// SIMATIC S7-200 SMART project (STEP 7-Micro/WIN SMART), CPU SR30

SYMBOL_TABLE STATES
RUNNING_STATE    M4.0     // RUNNING STATE
ON_STATE         M0.0     // ON STATE
PROCESS          M0.1     // PROCESS START
X_AXIS_STATE     M0.2     // X_AXIS_STATE
Y_AXIS_STATE     M0.3     // Y_AXIS_STATE
GRIPPER_STATE    M0.4     // GRIPPER_STATE
PROGRAM_STARTED  M0.5     // PROGRAM STARTED
READY_STATE      M0.6     // READY_STATE
PAUSE_STATE      M0.7     // PAUSE_STATE
END_SYMBOL_TABLE

SYMBOL_TABLE STEPS
STEP_1_DONE      M1.0     // STEP_1_DONE
STEP_2_DONE      M1.1     // STEP_2_DONE
STEP_3_DONE      M1.2     // STEP_3_DONE
STEP_4_DONE      M1.3     // STEP_4_DONE
STEP_5_DONE      M1.4     // STEP_5_DONE
STEP_6_DONE      M1.5     // STEP_6_DONE
STEP_7_DONE      M1.6     // STEP_7_DONE
STEP_8_DONE      M1.7     // STEP_8_DONE
END_SYMBOL_TABLE

SYMBOL_TABLE HMI INPUTSS
HMI_START        M2.0     // HMI_START
HMI_PAUSE        M2.1     // HMI_PAUSE
HMI_STOP         M2.2     // HMI_STOP
HMI_E_STOP       M2.3     // HMI_E_STOP
END_SYMBOL_TABLE

SYMBOL_TABLE MASTER INPUTS
MASTER_STOP      V202.5   // MASTER_STOP
MASTER_START     V201.5   // MASTER_START
MASTER_RESET     V203.5   // MASTER_RESET
COMMUNCATION     M6.0     // COMMUNCATION
END_SYMBOL_TABLE

ORGANIZATION_BLOCK MAIN:OB1
TITLE=Program Comments
BEGIN
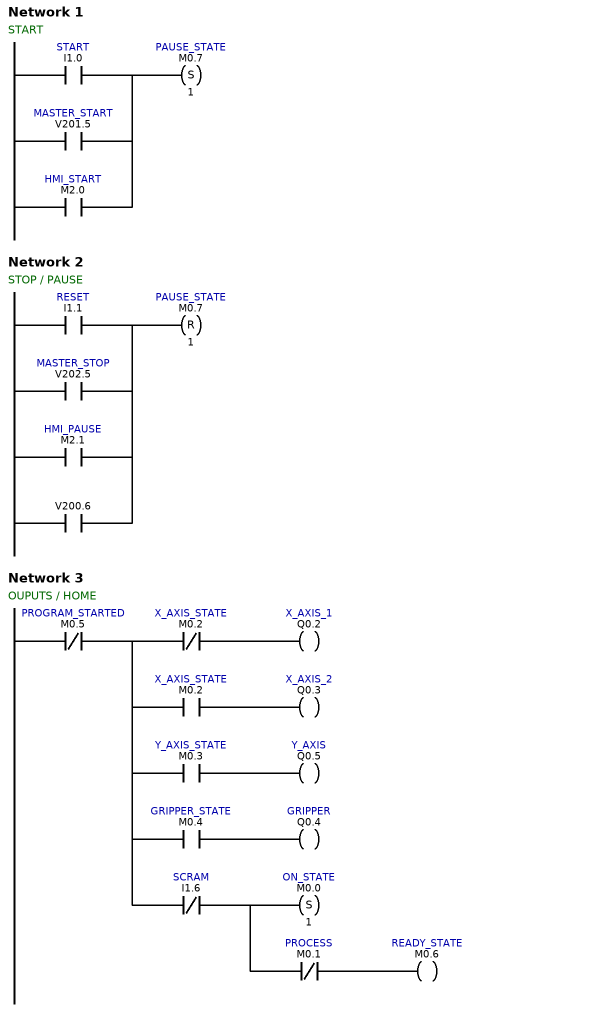
Network 1
// START
LD     START:I1.0
O      MASTER_START:V201.5
O      HMI_START:M2.0
S      PAUSE_STATE:M0.7, 1
Network 2
// STOP / PAUSE
LD     RESET:I1.1
O      MASTER_STOP:V202.5
O      HMI_PAUSE:M2.1
O      V200.6
R      PAUSE_STATE:M0.7, 1
Network 3
// OUPUTS / HOME
LDN    PROGRAM_STARTED:M0.5
LPS
AN     X_AXIS_STATE:M0.2
=      X_AXIS_1:Q0.2
LRD
A      X_AXIS_STATE:M0.2
=      X_AXIS_2:Q0.3
LRD
A      Y_AXIS_STATE:M0.3
=      Y_AXIS:Q0.5
LRD
A      GRIPPER_STATE:M0.4
=      GRIPPER:Q0.4
LPP
AN     SCRAM:I1.6
S      ON_STATE:M0.0, 1
AN     PROCESS:M0.1
=      READY_STATE:M0.6
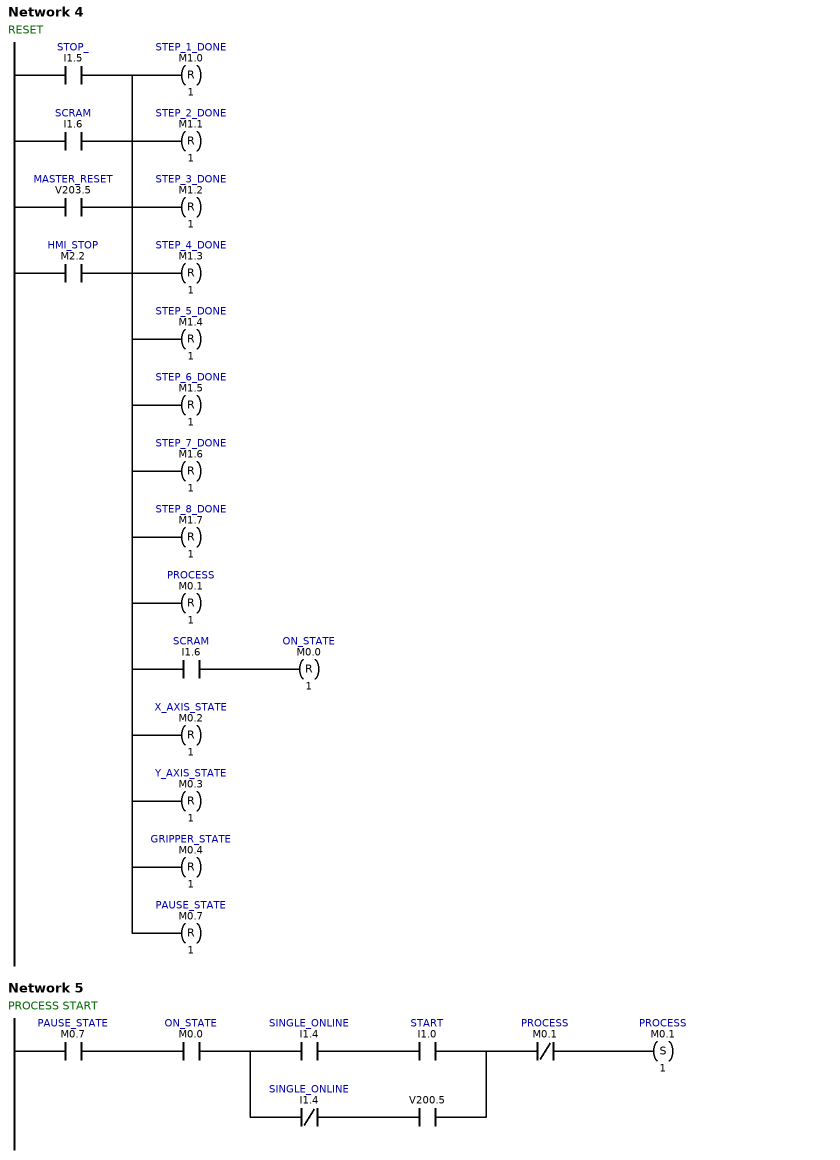
Network 4
// RESET 
LD     STOP_:I1.5
O      SCRAM:I1.6
O      MASTER_RESET:V203.5
O      HMI_STOP:M2.2
LPS
R      STEP_1_DONE:M1.0, 1
R      STEP_2_DONE:M1.1, 1
R      STEP_3_DONE:M1.2, 1
R      STEP_4_DONE:M1.3, 1
R      STEP_5_DONE:M1.4, 1
R      STEP_6_DONE:M1.5, 1
R      STEP_7_DONE:M1.6, 1
R      STEP_8_DONE:M1.7, 1
R      PROCESS:M0.1, 1
A      SCRAM:I1.6
R      ON_STATE:M0.0, 1
LRD
R      X_AXIS_STATE:M0.2, 1
LRD
R      Y_AXIS_STATE:M0.3, 1
LRD
R      GRIPPER_STATE:M0.4, 1
LPP
R      PAUSE_STATE:M0.7, 1
Network 5
// PROCESS START
LD     PAUSE_STATE:M0.7
A      ON_STATE:M0.0
LD     SINGLE_ONLINE:I1.4
A      START:I1.0
LDN    SINGLE_ONLINE:I1.4
A      V200.5
OLD
ALD
AN     PROCESS:M0.1
S      PROCESS:M0.1, 1
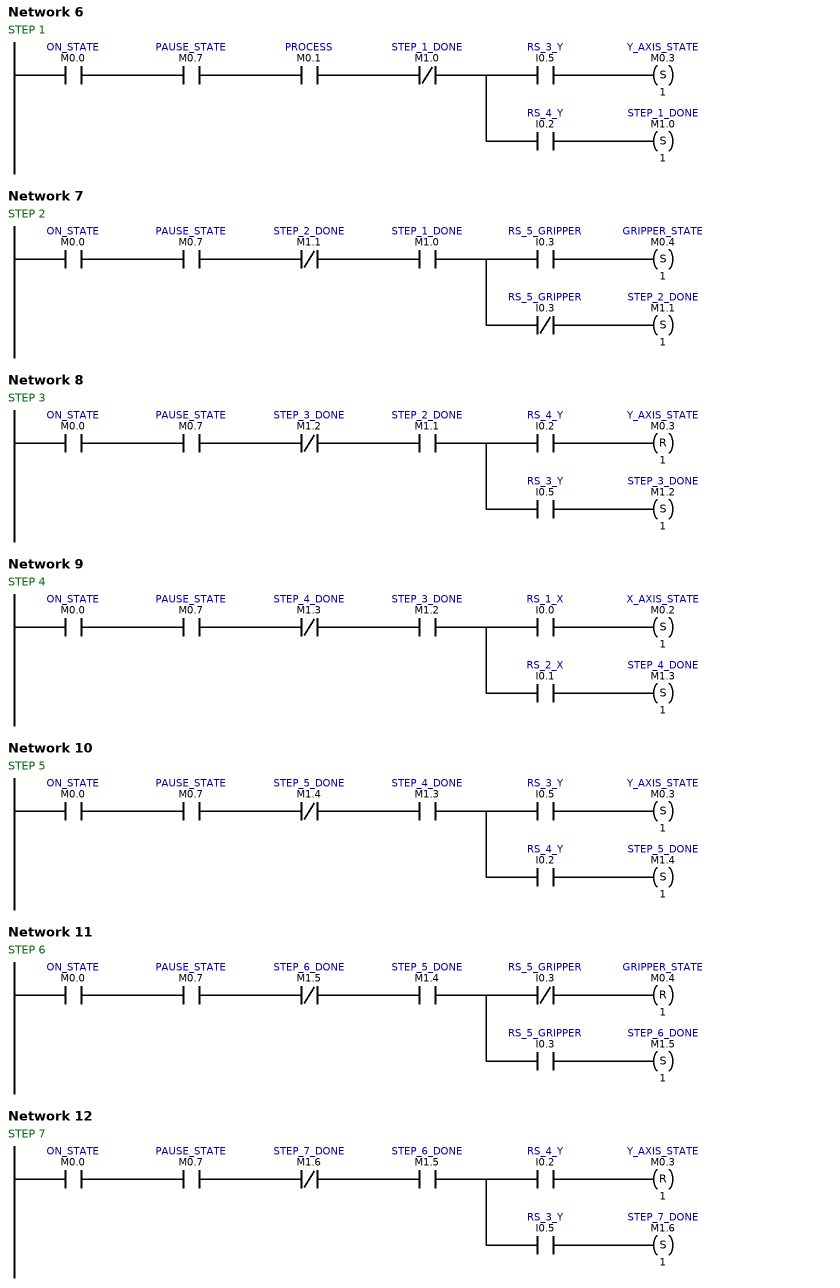
Network 6
// STEP 1
LD     ON_STATE:M0.0
A      PAUSE_STATE:M0.7
A      PROCESS:M0.1
AN     STEP_1_DONE:M1.0
LPS
A      RS_3_Y:I0.5
S      Y_AXIS_STATE:M0.3, 1
LPP
A      RS_4_Y:I0.2
S      STEP_1_DONE:M1.0, 1
Network 7
// STEP 2
LD     ON_STATE:M0.0
A      PAUSE_STATE:M0.7
AN     STEP_2_DONE:M1.1
A      STEP_1_DONE:M1.0
LPS
A      RS_5_GRIPPER:I0.3
S      GRIPPER_STATE:M0.4, 1
LPP
AN     RS_5_GRIPPER:I0.3
S      STEP_2_DONE:M1.1, 1
Network 8
// STEP 3
LD     ON_STATE:M0.0
A      PAUSE_STATE:M0.7
AN     STEP_3_DONE:M1.2
A      STEP_2_DONE:M1.1
LPS
A      RS_4_Y:I0.2
R      Y_AXIS_STATE:M0.3, 1
LPP
A      RS_3_Y:I0.5
S      STEP_3_DONE:M1.2, 1
Network 9
// STEP 4
LD     ON_STATE:M0.0
A      PAUSE_STATE:M0.7
AN     STEP_4_DONE:M1.3
A      STEP_3_DONE:M1.2
LPS
A      RS_1_X:I0.0
S      X_AXIS_STATE:M0.2, 1
LPP
A      RS_2_X:I0.1
S      STEP_4_DONE:M1.3, 1
Network 10
// STEP 5
LD     ON_STATE:M0.0
A      PAUSE_STATE:M0.7
AN     STEP_5_DONE:M1.4
A      STEP_4_DONE:M1.3
LPS
A      RS_3_Y:I0.5
S      Y_AXIS_STATE:M0.3, 1
LPP
A      RS_4_Y:I0.2
S      STEP_5_DONE:M1.4, 1
Network 11
// STEP 6
LD     ON_STATE:M0.0
A      PAUSE_STATE:M0.7
AN     STEP_6_DONE:M1.5
A      STEP_5_DONE:M1.4
LPS
AN     RS_5_GRIPPER:I0.3
R      GRIPPER_STATE:M0.4, 1
LPP
A      RS_5_GRIPPER:I0.3
S      STEP_6_DONE:M1.5, 1
Network 12
// STEP 7
LD     ON_STATE:M0.0
A      PAUSE_STATE:M0.7
AN     STEP_7_DONE:M1.6
A      STEP_6_DONE:M1.5
LPS
A      RS_4_Y:I0.2
R      Y_AXIS_STATE:M0.3, 1
LPP
A      RS_3_Y:I0.5
S      STEP_7_DONE:M1.6, 1
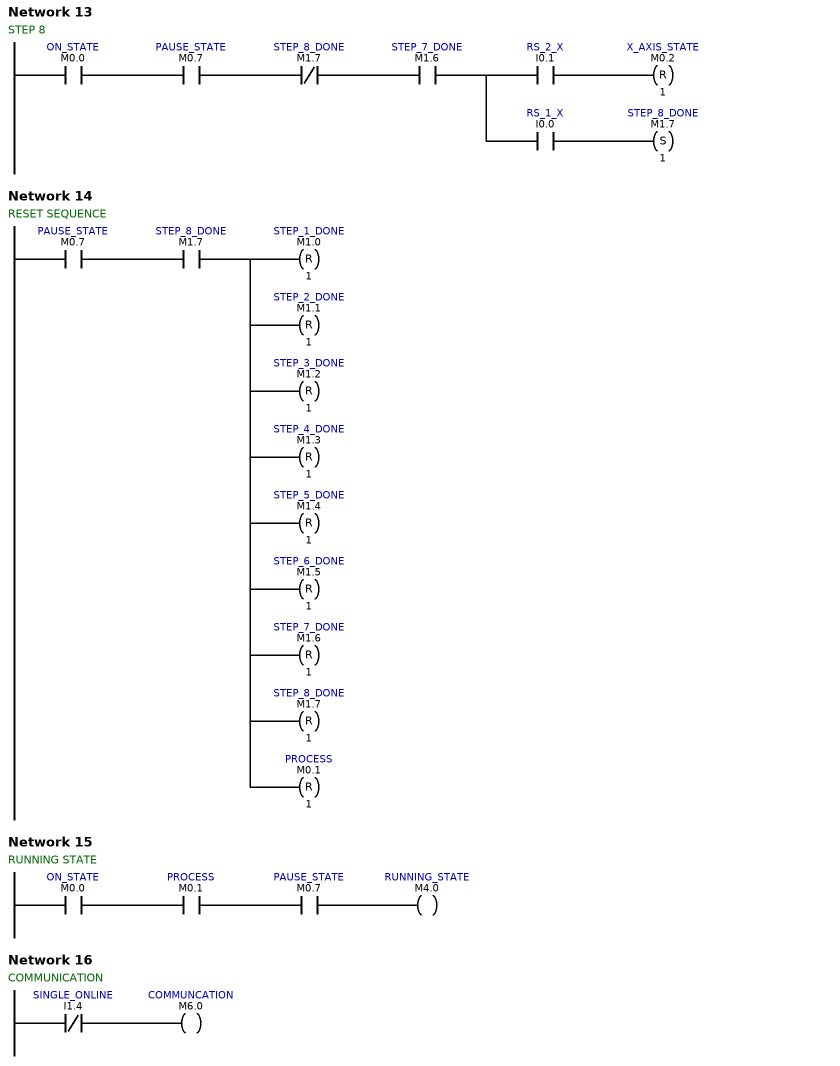
Network 13
// STEP 8
LD     ON_STATE:M0.0
A      PAUSE_STATE:M0.7
AN     STEP_8_DONE:M1.7
A      STEP_7_DONE:M1.6
LPS
A      RS_2_X:I0.1
R      X_AXIS_STATE:M0.2, 1
LPP
A      RS_1_X:I0.0
S      STEP_8_DONE:M1.7, 1
Network 14
// RESET SEQUENCE
LD     PAUSE_STATE:M0.7
A      STEP_8_DONE:M1.7
R      STEP_1_DONE:M1.0, 1
R      STEP_2_DONE:M1.1, 1
R      STEP_3_DONE:M1.2, 1
R      STEP_4_DONE:M1.3, 1
R      STEP_5_DONE:M1.4, 1
R      STEP_6_DONE:M1.5, 1
R      STEP_7_DONE:M1.6, 1
R      STEP_8_DONE:M1.7, 1
R      PROCESS:M0.1, 1
Network 15
// RUNNING STATE 
LD     ON_STATE:M0.0
A      PROCESS:M0.1
A      PAUSE_STATE:M0.7
=      RUNNING_STATE:M4.0
Network 16
// COMMUNICATION
LDN    SINGLE_ONLINE:I1.4
=      COMMUNCATION:M6.0
END_ORGANIZATION_BLOCK
